Fanuc KAREL source: kt00307.KL

-- PROVISIONAL review KL for V770-1; original PC SHA256 54b222aa1bea30b94089ee7f0603b65fb001073b3605ca80b49fea8fbe6c59cc
-- Incomplete behavior may be omitted. Consult companion uncertainty JSON. Do not deploy.
PROGRAM KT00307
%NOLOCKGROUP
VAR
  I2 : INTEGER
  OUT : BOOLEAN
-- UNRESOLVED_DECL H1 type=002017
BEGIN
  -- UNRESOLVED_PC offsets 5-19; opcodes 2E,22,9D,33,B4
  -- UNRESOLVED_PC offsets 24-35; opcodes 2E,23
  -- UNRESOLVED_PC offsets 40-62; opcodes 22,9D,33,B3,21,58,23
  -- UNRESOLVED_PC offsets 67-71; opcodes 7F
END KT00307
